// TIA Portal V19 export
// export: Created 2026-10-15T09:44:23.6112898Z, ExportSetting WithDefaults, DisplayName Totally Integrated Automation Portal, DisplayVersion V19, DisplayName TIA Portal Openness, DisplayVersion V19, DisplayName TIA Portal Version Control Interface, DisplayVersion V19, DisplayName STEP 7 Professional, DisplayVersion V19, DisplayName STEP 7 Safety, DisplayVersion V19, DisplayName WinCC Basic/Comfort/Advanced, DisplayVersion V19, DisplayName WinCC Unified, DisplayVersion V19
FUNCTION "ROLL_PB7" : Void   // FC17, SCL
{ S7_Optimized_Access := 'TRUE' }
VERSION : 0.1
// stored: AutoNumber true, IsIECCheckEnabled false, SetENOAutomatically false, UDAEnableTagReadback false
   VAR_TEMP
      r : Bool;
      a1 : Word;
      a2 : Word;
      activeDataBlock : Int;
      comparisonResults : Array[0..0] of Bool;
   END_VAR
BEGIN

   #r := FALSE;
   #a1 := W#16#0000;
   #a2 := W#16#0000;
   #activeDataBlock := 0;
   // PB7, STEP 5 network 1
   #r := ((NOT "ROLL_State".M[70, 2]) AND (NOT "ROLL_State".M[70, 3]) AND (NOT "ROLL_State".M[70, 4]) AND (NOT "ROLL_State".M[70, 6]) AND "ROLL_IO".Input[11, 0] AND "ROLL_IO".Input[11, 6] AND "ROLL_IO".Input[13, 3] AND "ROLL_State".M[63, 1]);
   "ROLL_State".M[28, 0] := #r;
   // PB7, STEP 5 network 2
   #r := ("ROLL_IO".Input[12, 1] AND "ROLL_IO".Input[12, 7]);
   "ROLL_State".M[28, 1] := #r;
   // PB7, STEP 5 network 3
   #r := ((NOT "ROLL_IO".Output[112, 5]) AND ((NOT "ROLL_IO".Output[112, 0]) OR (NOT "ROLL_State".M[31, 4])));
   "ROLL_State".M[28, 2] := #r;
   // PB7, STEP 5 network 4
   #r := (((NOT "ROLL_IO".Output[113, 0]) AND (NOT "ROLL_IO".Output[113, 1]) AND (NOT "ROLL_IO".Output[113, 3]) AND (NOT "ROLL_IO".Output[113, 5]) AND (NOT "ROLL_IO".Input[123, 5]) AND (NOT "ROLL_IO".Input[123, 6]) AND "ROLL_IO".Output[113, 2] AND "ROLL_IO".Output[113, 4] AND "ROLL_IO".Input[124, 1] AND "ROLL_IO".Input[124, 4]) OR "ROLL_State".M[0, 4]);
   "ROLL_State".M[240, 0] := #r;
   // PB7, STEP 5 network 5
   #r := ((((NOT "ROLL_IO".Output[113, 2]) AND "ROLL_IO".Output[113, 3] AND "ROLL_IO".Input[123, 5] AND "ROLL_IO".Input[124, 1] AND "ROLL_IO".Input[124, 4]) OR ((NOT "ROLL_IO".Output[113, 3]) AND "ROLL_IO".Output[113, 2] AND "ROLL_IO".Input[124, 1] AND "ROLL_IO".Input[124, 5]) OR "ROLL_State".M[0, 4]) AND "ROLL_State".M[20, 2]);
   "ROLL_State".M[240, 1] := #r;
   // PB7, STEP 5 network 6
   #r := ("ROLL_State".M[240, 0] OR "ROLL_State".M[240, 1]);
   "ROLL_State".M[28, 3] := #r;
   // PB7, STEP 5 network 7
   #r := ("ROLL_State".M[28, 0] AND "ROLL_State".M[28, 1] AND "ROLL_State".M[28, 2] AND "ROLL_State".M[28, 3]);
   "ROLL_State".M[28, 4] := #r;
   // PB7, STEP 5 network 8
   #r := ("ROLL_IO".Input[10, 7] AND "ROLL_IO".Input[3, 4] AND "ROLL_IO".Input[3, 5] AND "ROLL_IO".Input[3, 7]);
   "ROLL_State".M[28, 5] := #r;
   // PB7, STEP 5 network 9
   #r := ((NOT "ROLL_State".M[13, 4]) AND (NOT "ROLL_State".M[16, 6]) AND (NOT "ROLL_State".M[5, 7]) AND "ROLL_State".M[28, 5]);
   "ROLL_State".M[28, 6] := #r;
   // PB7, STEP 5 network 10
   #r := (("ROLL_IO".Input[0, 2] AND "ROLL_IO".Input[0, 4]) OR "ROLL_IO".Input[0, 1]);
   IF #r THEN
       "ROLL_State".M[29, 0] := TRUE;
   END_IF;
   #r := (NOT "ROLL_State".M[28, 6]);
   IF #r THEN
       "ROLL_State".M[29, 0] := FALSE;
   END_IF;
   // PB7, STEP 5 network 11
   #r := ("ROLL_State".M[29, 0] AND "ROLL_State".S5Timers[13].Q);
   "ROLL_State".M[29, 1] := #r;
   // PB7, STEP 5 network 12
   #r := (NOT "ROLL_State".M[12, 1]);
   "ROLL_State".M[30, 0] := #r;
   // PB7, STEP 5 network 13
   #r := "ROLL_State".M[0, 4];
   "ROLL_State".M[30, 1] := #r;
   // PB7, STEP 5 network 14
   #r := ((NOT "ROLL_State".M[6, 1]) AND (NOT "ROLL_State".M[6, 3]) AND (NOT "ROLL_State".M[6, 4]) AND (NOT "ROLL_State".M[6, 5]) AND (NOT "ROLL_State".M[6, 6]) AND (NOT "ROLL_State".M[6, 7]) AND (NOT "ROLL_State".M[7, 0]) AND (NOT "ROLL_State".M[7, 1]) AND (NOT "ROLL_State".M[7, 2]) AND (NOT "ROLL_State".M[7, 3]) AND (NOT "ROLL_State".M[7, 7]));
   "ROLL_State".M[30, 2] := #r;
   // PB7, STEP 5 network 15
   #r := ((NOT "ROLL_IO".Input[3, 6]) AND (NOT "ROLL_State".M[5, 6]));
   "ROLL_State".M[30, 3] := #r;
   // PB7, STEP 5 network 16
   #r := (("ROLL_State".M[30, 0] AND "ROLL_State".M[30, 1] AND "ROLL_State".M[30, 2] AND "ROLL_State".M[30, 3]) OR "ROLL_IO".Input[0, 0] OR "ROLL_IO".Input[0, 6]);
   "ROLL_State".M[30, 5] := #r;
   // PB7, STEP 5 network 17
   #r := ((NOT "ROLL_State".M[11, 0]) AND (NOT "ROLL_State".M[13, 1]) AND (NOT "ROLL_State".M[13, 3]) AND (NOT "ROLL_State".M[5, 0]) AND (NOT "ROLL_State".M[5, 1]) AND (NOT "ROLL_State".M[5, 2]));
   "ROLL_State".M[30, 6] := #r;
   // PB7, STEP 5 network 18
   #r := ((NOT "ROLL_State".M[11, 1]) AND (NOT "ROLL_State".M[5, 3]) AND (NOT "ROLL_State".M[9, 1]) AND (NOT "ROLL_State".M[9, 2]) AND (NOT "ROLL_State".M[9, 3]) AND "ROLL_IO".Input[8, 5] AND "ROLL_State".M[28, 6]);
   "ROLL_State".M[30, 7] := #r;
   // PB7, STEP 5 network 19
   #r := ((NOT "ROLL_State".M[12, 0]) AND (NOT "ROLL_State".M[9, 0]));
   "ROLL_State".M[31, 0] := #r;
   // PB7, STEP 5 network 20
   #r := ((NOT "ROLL_State".M[87, 5]) AND (NOT "ROLL_State".M[88, 1]) AND (NOT "ROLL_State".M[88, 3]) AND (NOT "ROLL_State".M[88, 4]) AND (NOT "ROLL_State".M[88, 5]) AND (NOT "ROLL_State".M[88, 6]));
   "ROLL_State".M[31, 2] := #r;
   // PB7, STEP 5 network 21
   #r := ("ROLL_State".M[30, 5] AND "ROLL_State".M[30, 6] AND "ROLL_State".M[30, 7] AND "ROLL_State".M[31, 0] AND "ROLL_State".M[31, 2]);
   "ROLL_State".M[31, 1] := #r;
   // PB7, STEP 5 network 22
   #r := (("ROLL_State".M[28, 4] OR "ROLL_State".M[31, 5]) AND "ROLL_IO".Input[0, 4] AND "ROLL_State".M[4, 4]);
   IF #r THEN
       "ROLL_State".M[31, 4] := TRUE;
   END_IF;
   #r := ((NOT "ROLL_IO".Input[0, 2]) OR (NOT "ROLL_IO".Input[0, 3]) OR (NOT "ROLL_State".M[29, 0]) OR (NOT "ROLL_State".M[31, 1]));
   IF #r THEN
       "ROLL_State".M[31, 4] := FALSE;
   END_IF;
   // PB7, STEP 5 network 23
   #r := "ROLL_State".M[31, 4];
   IF #r THEN
       "ROLL_State".M[31, 5] := TRUE;
   END_IF;
   #r := (((NOT "ROLL_State".M[31, 4]) AND (((NOT "ROLL_State".M[37, 2]) AND "ROLL_State".M[37, 1]) OR "ROLL_State".M[37, 0]) AND "ROLL_State".M[28, 4]) OR (NOT "ROLL_IO".Input[0, 2]));
   IF #r THEN
       "ROLL_State".M[31, 5] := FALSE;
   END_IF;
   // PB7, STEP 5 network 24
   #r := "ROLL_State".M[52, 3];
   IF #r THEN
       "ROLL_State".M[31, 6] := TRUE;
   END_IF;
   #r := ((NOT "ROLL_IO".Input[14, 0]) AND "ROLL_IO".Input[12, 1]);
   IF #r THEN
       "ROLL_State".M[31, 6] := FALSE;
   END_IF;
   // PB7, STEP 5 network 25
   #r := "ROLL_State".M[31, 5];
   "ROLL_IO".Output[16, 6] := #r;
   // PB7, STEP 5 network 26
   #r := "ROLL_State".M[40, 0];
   "ROLL_IO".Output[16, 7] := #r;
   // PB7, STEP 5 network 27
   RETURN;
END_FUNCTION
